Omron CX-Programmer project NewProject (CX-Programmer 9.75)

# PLC Flicker_Operation_Timer: CP1E N30

## Global symbols (name address type ; comment)
0.00 BOOL  ; SW1 (X24)
100.00 BOOL  ; Y1
T000 BOOL  ; T3
T001 BOOL  ; T4

## Program NewProgram1 (cyclic task 0)

### Section Section1

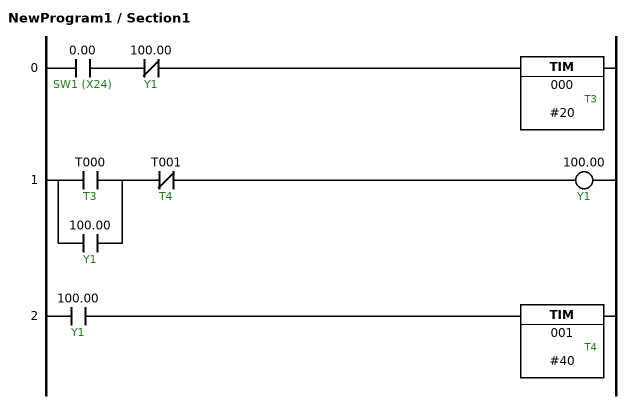
; rung 0
LD 0.00  ; SW1 (X24)
ANDNOT 100.00  ; Y1
TIM 000 #20  ; T3
; rung 1
LD T000  ; T3
OR 100.00  ; Y1
ANDNOT T001  ; T4
OUT 100.00  ; Y1
; rung 2
LD 100.00  ; Y1
TIM 001 #40  ; T4

### Section END
; rung 0
END(001)